Universal Robots URScript: T010_qwen2.5-coder_32b_baseline_rep3.urscript

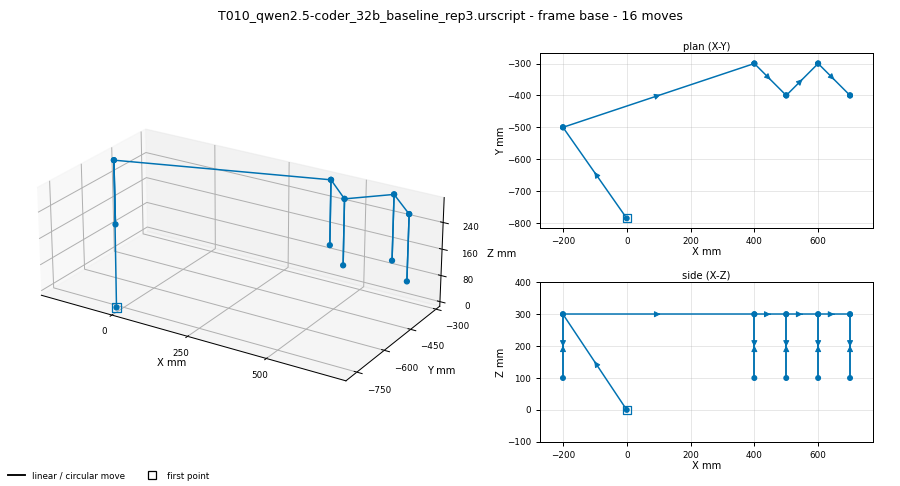
[picture p0: tool path of T010_qwen2.5-coder_32b_baseline_rep3.urscript in frame base, 16 of 16 moves have a stored position in this frame; points joined in program order, loops and branches not executed]
# Move to Home position
movej(p[0.0, -0.7854, 0.0, -2.3562, -1.5708, 0.0], a=1.4, v=1.05)

# Move above screw feeder
movel(p[-0.2, -0.5, 0.3, -2.3562, -1.5708, 0.0], a=1.2, v=1.05)

# Pick screw from feeder
movel(p[-0.2, -0.5, 0.1, -2.3562, -1.5708, 0.0], a=1.2, v=0.4)

# Lift from feeder
movel(p[-0.2, -0.5, 0.3, -2.3562, -1.5708, 0.0], a=1.2, v=0.9)

# Move above fastening point 1
movel(p[0.4, -0.3, 0.3, -2.3562, -1.5708, 0.0], a=1.2, v=1.05)

# Fasten at point 1 (fenced mode)
set_tcp(p[-0.004, 0.004, 0.1, 3.1416, -0.7854, 0])
movel(p[0.4, -0.3, 0.1, -2.3562, -1.5708, 0.0], a=0.5, v=0.2)
sleep(1) # Simulate fastening time
movel(p[0.4, -0.3, 0.3, -2.3562, -1.5708, 0.0], a=0.5, v=0.9)

# Move above fastening point 2
movel(p[0.5, -0.4, 0.3, -2.3562, -1.5708, 0.0], a=1.2, v=1.05)

# Fasten at point 2 (fenced mode)
movel(p[0.5, -0.4, 0.1, -2.3562, -1.5708, 0.0], a=0.5, v=0.2)
sleep(1) # Simulate fastening time
movel(p[0.5, -0.4, 0.3, -2.3562, -1.5708, 0.0], a=0.5, v=0.9)

# Move above fastening point 3
movel(p[0.6, -0.3, 0.3, -2.3562, -1.5708, 0.0], a=1.2, v=1.05)

# Fasten at point 3 (fenced mode)
movel(p[0.6, -0.3, 0.1, -2.3562, -1.5708, 0.0], a=0.5, v=0.2)
sleep(1) # Simulate fastening time
movel(p[0.6, -0.3, 0.3, -2.3562, -1.5708, 0.0], a=0.5, v=0.9)

# Move above fastening point 4
movel(p[0.7, -0.4, 0.3, -2.3562, -1.5708, 0.0], a=1.2, v=1.05)

# Fasten at point 4 (fenced mode)
movel(p[0.7, -0.4, 0.1, -2.3562, -1.5708, 0.0], a=0.5, v=0.2)
sleep(1) # Simulate fastening time
movel(p[0.7, -0.4, 0.3, -2.3562, -1.5708, 0.0], a=0.5, v=0.9)

# Reset TCP to default
set_tcp(p[0.0, 0.0, 0.0, 0.0, 0.0, 0.0])
